// TIA Portal V20 export
// export: Created 2026-10-19T18:06:14.0811462Z, ExportSetting WithDefaults, DisplayName Totally Integrated Automation Portal, DisplayVersion V20 Update 6, DisplayName TIA Portal Openness, DisplayVersion V20 Update 6, DisplayName TIA Portal Version Control Interface, DisplayVersion V20 Update 6, DisplayName SINAMICS Startdrive Advanced, DisplayVersion V20 SP1, DisplayName SINAMICS Startdrive G130, G150, S120, S150, SINAMICS MV, G220, S200, S210, DisplayVersion V20 SP1, DisplayName SINAMICS Startdrive G110M, G120, G120C, G120D, G120P, G115D, DisplayVersion V20 SP1, DisplayName STEP 7 Professional, DisplayVersion V20 Update 6, DisplayName STEP 7 Safety, DisplayVersion V20 Update 2, DisplayName WinCC Basic/Comfort/Advanced, DisplayVersion V20 Update 6, DisplayName WinCC Unified, DisplayVersion V20 Update 6
FUNCTION "SAI_Copy" : Void   // FC29, LAD
{ S7_Optimized_Access := 'FALSE' }
VERSION : 0.1
// stored: AutoNumber true, IsIECCheckEnabled false, SetENOAutomatically false, UDAEnableTagReadback false
   VAR_INPUT
      Src : Variant;
   END_VAR
   VAR_IN_OUT
      Dest : Variant;
   END_VAR
   VAR_TEMP
      TmpBuf : Array[0..100] of Byte;
      TmpRet : Int;
      TmpPos : DInt;
   END_VAR
BEGIN

REGION Network 1
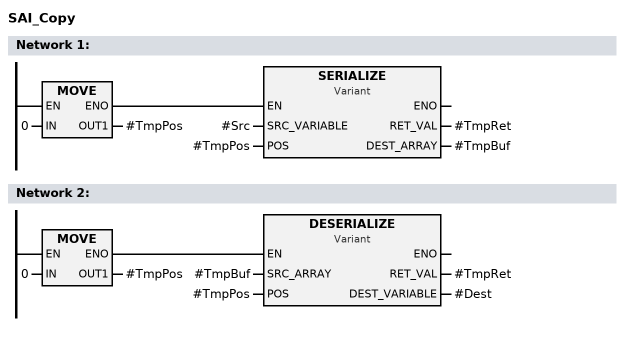
   RUNG wire#powerrail
      Move(in := 0, out1 => #TmpPos)
      { S7_Templates := "[src_type := Variant, dest_type := Variant]" } Serialize(SRC_VARIABLE := #Src, POS := #TmpPos, Ret_Val => #TmpRet, DEST_ARRAY => #TmpBuf)
   END_RUNG
   // the same network as SCL:
   #TmpPos := 0;
   #TmpRet := Serialize(SRC_VARIABLE := #Src, POS := #TmpPos, DEST_ARRAY => #TmpBuf);
END_REGION

REGION Network 2
   RUNG wire#powerrail
      Move(in := 0, out1 => #TmpPos)
      { S7_Templates := "[src_type := Variant, dest_type := Variant]" } Deserialize(SRC_ARRAY := #TmpBuf, POS := #TmpPos, Ret_Val => #TmpRet, DEST_VARIABLE => #Dest)
   END_RUNG
   // the same network as SCL:
   #TmpPos := 0;
   #TmpRet := Deserialize(SRC_ARRAY := #TmpBuf, POS := #TmpPos, DEST_VARIABLE => #Dest);
END_REGION
END_FUNCTION
